SYSTEM ResourceDeploymentTest
  (* Version 1.0, 2024-08-21, mario *)
  APPLICATION ResourceDeploymentTestApp
  END_APPLICATION
  DEVICE FORTE_PC : FORTE_PC(MGR_ID := "localhost:61499" (* Device manager socket ID *))
    {SET_ATTRIBUTE(Profile, HOLOBLOC)}
    RESOURCE TestNetwork_Empty : EMB_RES
    END_RESOURCE
    RESOURCE TestNetwork_StackedTypedSubapp : EMB_RES
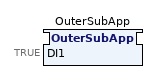
      SUBAPPS
        OuterSubApp : OuterSubApp(DI1 := TRUE);
      END_SUBAPPS
    END_RESOURCE
    RESOURCE TestNetwork_StackedUntypedSubapp : EMB_RES
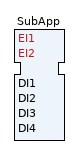
      SUBAPPLICATION SubApp
        EVENT_INPUT
          EI1;
          EI2;
        END_EVENT
        VAR_INPUT
          DI1 : INT;
          DI2 : BOOL;
          DI3 : STRING;
          DI4 : BOOL := TRUE;
        END_VAR
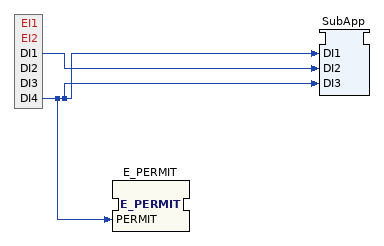
        FBS
          E_PERMIT : E_PERMIT;
        END_FBS
        SUBAPPLICATION SubApp
          VAR_INPUT
            DI1 : BOOL;
            DI2 : INT;
            DI3 : BOOL;
          END_VAR
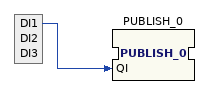
          FBS
            PUBLISH_0 : PUBLISH_0;
          END_FBS
          DATA_CONNECTIONS
            DI1 TO PUBLISH_0.QI;
          END_CONNECTIONS
        END_SUBAPPLICATION
        DATA_CONNECTIONS
          DI4 TO E_PERMIT.PERMIT;
          DI4 TO SubApp.DI3;
          DI4 TO SubApp.DI1;
          DI1 TO SubApp.DI2;
        END_CONNECTIONS
      END_SUBAPPLICATION
    END_RESOURCE
  END_DEVICE
END_SYSTEM
